(* IEC 61131-3 sources: plcassist-cli/packages/volt-lsp-iec/test-corpus/lenze-mid/Device/Plc Logic/Application/Library Manager/(unresolved)/visu interfaces, 13 files *)

(* ---- GVL.gvl ---- *)
VAR_GLOBAL
	G_VISUCOMMANDMANAGER : ICommandManager;
	G_VISUCOMMANDMANAGER2 : ICommandManager2;
	G_GLOBALCLIENTMANAGER : IVisuGlobalClientManager;
END_VAR

(* ---- GVL_CONSTANT.gvl ---- *)
VAR_GLOBAL
	VISU_INVALID_ID : INT := -1;
END_VAR

(* ---- IATTACHEDVISUALELEMENT.itf ---- *)
INTERFACE IATTACHEDVISUALELEMENT
END_INTERFACE

METHOD GETLOCATION : VisuStructSimpleRectangleItf
END_METHOD

(* ---- IBUTTONCLIENTSTATE.itf ---- *)
INTERFACE IBUTTONCLIENTSTATE
END_INTERFACE

METHOD ISPRESSED : BOOL
END_METHOD

METHOD SETPRESSED
VAR_INPUT
	BPRESSED : BOOL;
END_VAR
END_METHOD

(* ---- ICOMMANDMANAGER.itf ---- *)
INTERFACE ICOMMANDMANAGER
END_INTERFACE

METHOD GETCOMMAND : IGeneralCommand
VAR_INPUT
	IINDEX : INT;
END_VAR
END_METHOD

METHOD REGISTERCOMMAND : BOOL
VAR_INPUT
	CMD : IGeneralCommand;
END_VAR
END_METHOD

METHOD UNREGISTERCOMMAND : BOOL
VAR_INPUT
	CMD : IGeneralCommand;
END_VAR
END_METHOD

(* ---- ICOMMANDMANAGER2.itf ---- *)
INTERFACE ICOMMANDMANAGER2
END_INTERFACE

METHOD GETCOMMAND : IGeneralCommand2
VAR_INPUT
	IINDEX : INT;
END_VAR
END_METHOD

METHOD REGISTERCOMMAND : BOOL
VAR_INPUT
	CMD : IGeneralCommand2;
END_VAR
END_METHOD

METHOD UNREGISTERCOMMAND : BOOL
VAR_INPUT
	CMD : IGeneralCommand2;
END_VAR
END_METHOD

(* ---- IGENERALCOMMAND.itf ---- *)
INTERFACE IGENERALCOMMAND
END_INTERFACE

METHOD EXECUTE : DWORD
VAR_INPUT
	DWPARAM1 : DWORD;
	DWPARAM2 : DWORD;
END_VAR
END_METHOD

(* ---- IGENERALCOMMAND2.itf ---- *)
INTERFACE IGENERALCOMMAND2
END_INTERFACE

METHOD EXECUTE : __XWORD
VAR_INPUT
	DWPARAM1 : __XWORD;
	DWPARAM2 : __XWORD;
END_VAR
END_METHOD

(* ---- IGENERIC.itf ---- *)
INTERFACE IGENERIC
END_INTERFACE

METHOD GETINTERFACE : POINTER TO BYTE
VAR_INPUT
	DWITFID : DWORD;
END_VAR
END_METHOD

(* ---- IGLOBALCLIENTMANAGERLISTENER.itf ---- *)
INTERFACE IGLOBALCLIENTMANAGERLISTENER
END_INTERFACE

METHOD CLIENTCREATED
VAR_INPUT
	IGLOBALCLIENTID : INT;
	EVISUCLIENTTYPE : Visu_ClientTypeItf;
END_VAR
END_METHOD

METHOD CLIENTDESTROYED
VAR_INPUT
	IGLOBALCLIENTID : INT;
	EVISUCLIENTTYPE : Visu_ClientTypeItf;
END_VAR
END_METHOD

(* ---- IVISUGLOBALCLIENTMANAGER.itf ---- *)
INTERFACE IVISUGLOBALCLIENTMANAGER
END_INTERFACE

METHOD REGISTERORUPDATECLIENT : INT
VAR_INPUT
	IGLOBALCLIENTID : INT;
	EVISUCLIENTTYPE : Visu_ClientTypeItf;
END_VAR
END_METHOD

METHOD SETCURRENTCLIENTID : BOOL
VAR_INPUT
	IGLOBALCLIENTID : INT;
END_VAR
END_METHOD

(* ---- IVISUGLOBALCLIENTMANAGER2.itf ---- *)
INTERFACE IVISUGLOBALCLIENTMANAGER2
END_INTERFACE

METHOD ADDGLOBALCLIENTMANAGERLISTENER : BOOL
VAR_INPUT
	ITFGLOBALCLIENTMANAGERLISTENER : IGlobalClientManagerListener;
END_VAR
END_METHOD

(* ---- IVISUGLOBALCLIENTMANAGER3.itf ---- *)
INTERFACE IVISUGLOBALCLIENTMANAGER3
END_INTERFACE

METHOD UNREGISTERCLIENT : BOOL
VAR_INPUT
	IGLOBALCLIENTID : INT;
	EVISUCLIENTTYPE : Visu_ClientTypeItf;
END_VAR
END_METHOD
